(* IEC 61131-3 sources: rusty/tests/lit/multi/external_unit_linkage/chain/lib_a, 7 files *)

(* ---- IBase.st ---- *)
INTERFACE IBase
    METHOD base_id : DINT END_METHOD
END_INTERFACE

(* ---- IShape.st ---- *)
INTERFACE IShape
    METHOD area : DINT
    VAR_INPUT
        unit : STRING[10];
    END_VAR
    END_METHOD
END_INTERFACE

(* ---- AbstractShape.st ---- *)
FUNCTION_BLOCK ABSTRACT AbstractShape IMPLEMENTS IShape
VAR_OUTPUT
    unit_seen : STRING[10];
END_VAR
    METHOD ABSTRACT area : DINT
    VAR_INPUT
        unit : STRING[10];
    END_VAR
    END_METHOD
END_FUNCTION_BLOCK

(* ---- Base.st ---- *)
FUNCTION_BLOCK Base IMPLEMENTS IBase
    METHOD base_id : DINT
        base_id := 1;
    END_METHOD

    METHOD kind : DINT
        kind := 10;
    END_METHOD
END_FUNCTION_BLOCK

(* ---- CBase.st ---- *)
CLASS CBase
    METHOD value : DINT
        value := 100;
    END_METHOD
END_CLASS

(* ---- Plain.st ---- *)
FUNCTION_BLOCK Plain
VAR_INPUT
    x : DINT := 2;
END_VAR
END_FUNCTION_BLOCK

(* ---- PropBase.st ---- *)
FUNCTION_BLOCK PropBase
VAR
    text : STRING[20] := 'base';
END_VAR
    PROPERTY_GET name : STRING[20]
        name := text;
    END_PROPERTY
END_FUNCTION_BLOCK
